Staubli VAL3: copyPara.pgx

public program copyPara(string x_sTarget, num x_nSource, num x_nTarget)
  local num l_nSize
  local num l_i
  local num l_j
begin

  progTemp:pProgItem[x_sTarget].pProgTemplate[x_nTarget].sTRAJname=progTemp:pProgItem[x_sTarget].pProgTemplate[x_nSource].sTRAJname
  progTemp:pProgItem[x_sTarget].pProgTemplate[x_nTarget].nType=progTemp:pProgItem[x_sTarget].pProgTemplate[x_nSource].nType
  for l_j=0 to 2
    progTemp:pProgItem[x_sTarget].pProgTemplate[x_nTarget].iIfItem.nSigType[l_j]=progTemp:pProgItem[x_sTarget].pProgTemplate[x_nSource].iIfItem.nSigType[l_j]
    progTemp:pProgItem[x_sTarget].pProgTemplate[x_nTarget].iIfItem.nSigIndex[l_j]=progTemp:pProgItem[x_sTarget].pProgTemplate[x_nSource].iIfItem.nSigIndex[l_j]
    progTemp:pProgItem[x_sTarget].pProgTemplate[x_nTarget].iIfItem.nValue[l_j]=progTemp:pProgItem[x_sTarget].pProgTemplate[x_nSource].iIfItem.nValue[l_j]
  endFor
  progTemp:pProgItem[x_sTarget].pProgTemplate[x_nTarget].iIfItem.bANDOR[0]=(progTemp:pProgItem[x_sTarget].pProgTemplate[x_nSource].iIfItem.bANDOR[0]==true)
  progTemp:pProgItem[x_sTarget].pProgTemplate[x_nTarget].iIfItem.bANDOR[1]=(progTemp:pProgItem[x_sTarget].pProgTemplate[x_nSource].iIfItem.bANDOR[1]==true)

end
